	mF_Mpc_b_Ac: ARRAY[0..731] OF LREAL := [-0.00028473180920350741, -0.00064838280152378558, -0.0010871186383875045, -0.0015972149310527575, -0.0021750553811336337, -0.0028171299154482626, -0.0035200328169797839, -0.00428046085366274, -0.0050952114066324721, -0.0059611805995021831, -0.0068753614301614151, -0.0078348419065206853, -0.00883680318755997, -0.0098785177309735454, -0.010957347448640358, -0.012070741871087625, -0.013216236322055611, -0.014391450104213641, -0.015594084697021157, -0.016821921967673122, -0.018072822396016243, -0.019344723314271256, -0.02063563716234695, -0.021943649759483548, -0.023266918592916585, -0.024603671124207489, -0.025952203113843546, -0.027310876964667902, -0.02867812008465969, -0.030052423269545051, -0.031432339105682078, -0.032816480393626085, -0.034203518592746424, -0.035592182287232092, -0.036981255673790715, -0.038369577071313908, -0.039756037452751761, -0.041139578999410086, -0.042519193677855886, -0.043893921839589789, -0.04526285084361819, -0.046625113702033094, -0.047979887748683912, -0.049326393331002638, -0.050663892525022049, -0.051991687873605683, -0.053309121147888459, -0.054615572131907646, -0.055910457430385821, -0.057193229299610078, -0.058463374501335187, -0.05972041317962274, -0.06096389776051344, -0.062193411874415308, -0.063408569301077411, -0.0646090129370057, -0.065794413785165692, -0.066964469966805218, -0.068118905755219825, -0.069257470631273188, -0.070379938360475486, -0.071486106091413787, -0.072575793475319991, -0.073648841806554288, -0.074705113183774638, -0.075744489691556227, -0.076766872602218345, -0.077772181597610637, -0.078760354010605146, -0.079731344086035758, -0.080685122260822376, -0.081621674463012911, -0.082541001429472627, -0.08344311804194729, -0.084328052681223467, -0.085195846599106978, -0.086046553307938353, -0.08688023798736208, -0.087696976908065286, -0.088496856872199881, -0.089279974670201517, -0.090046436553718037, -0.0907963577243595, -0.091529861837982063, -0.092247080524217845, -0.0929481529209633, -0.093633225223539271, -0.094302450248236622, -0.094955987009962314, -0.0955940003137019, -0.096216660359515871, -0.096824142360788817, -0.09741662617545184, -0.0979942959499008, -0.098557339775334651, -0.099105949356240508, -0.099640319690754223, -0.10016064876262748, -0.1006671372445353, -0.10115998821245992, -0.10163940687089022, -0.10210560028857829, -0.10255877714459775, -0.10299914748445149, -0.10342692248597933, -0.10384231423481935, -0.10424553550917975, -0.10463679957368147, -0.10501631998203463, -0.105384310388316, -0.10574098436661702, -0.10608655523883639, -0.10642123591039374, -0.10674523871364502, -0.10705877525878353, -0.1073620562920138, -0.1076552915607895, -0.10793868968590982, -0.10821245804027231, -0.10847680263408387, 0.00028473180920350741, 0.00064838280152378558, 0.0010871186383875045, 0.0015972149310527575, 0.0021750553811336337, 0.0028171299154482626, 0.0035200328169797839, 0.00428046085366274, 0.0050952114066324721, 0.0059611805995021831, 0.0068753614301614151, 0.0078348419065206853, 0.00883680318755997, 0.0098785177309735454, 0.010957347448640358, 0.012070741871087625, 0.013216236322055611, 0.014391450104213641, 0.015594084697021157, 0.016821921967673122, 0.018072822396016243, 0.019344723314271256, 0.02063563716234695, 0.021943649759483548, 0.023266918592916585, 0.024603671124207489, 0.025952203113843546, 0.027310876964667902, 0.02867812008465969, 0.030052423269545051, 0.031432339105682078, 0.032816480393626085, 0.034203518592746424, 0.035592182287232092, 0.036981255673790715, 0.038369577071313908, 0.039756037452751761, 0.041139578999410086, 0.042519193677855886, 0.043893921839589789, 0.04526285084361819, 0.046625113702033094, 0.047979887748683912, 0.049326393331002638, 0.050663892525022049, 0.051991687873605683, 0.053309121147888459, 0.054615572131907646, 0.055910457430385821, 0.057193229299610078, 0.058463374501335187, 0.05972041317962274, 0.06096389776051344, 0.062193411874415308, 0.063408569301077411, 0.0646090129370057, 0.065794413785165692, 0.066964469966805218, 0.068118905755219825, 0.069257470631273188, 0.070379938360475486, 0.071486106091413787, 0.072575793475319991, 0.073648841806554288, 0.074705113183774638, 0.075744489691556227, 0.076766872602218345, 0.077772181597610637, 0.078760354010605146, 0.079731344086035758, 0.080685122260822376, 0.081621674463012911, 0.082541001429472627, 0.08344311804194729, 0.084328052681223467, 0.085195846599106978, 0.086046553307938353, 0.08688023798736208, 0.087696976908065286, 0.088496856872199881, 0.089279974670201517, 0.090046436553718037, 0.0907963577243595, 0.091529861837982063, 0.092247080524217845, 0.0929481529209633, 0.093633225223539271, 0.094302450248236622, 0.094955987009962314, 0.0955940003137019, 0.096216660359515871, 0.096824142360788817, 0.09741662617545184, 0.0979942959499008, 0.098557339775334651, 0.099105949356240508, 0.099640319690754223, 0.10016064876262748, 0.1006671372445353, 0.10115998821245992, 0.10163940687089022, 0.10210560028857829, 0.10255877714459775, 0.10299914748445149, 0.10342692248597933, 0.10384231423481935, 0.10424553550917975, 0.10463679957368147, 0.10501631998203463, 0.105384310388316, 0.10574098436661702, 0.10608655523883639, 0.10642123591039374, 0.10674523871364502, 0.10705877525878353, 0.1073620562920138, 0.1076552915607895, 0.10793868968590982, 0.10821245804027231, 0.10847680263408387, -1.0, -1.0, 1.0, 1.0, -0.0, -0.00028473180920350741, -0.00064838280152378558, -0.0010871186383875045, -0.0015972149310527575, -0.0021750553811336337, -0.0028171299154482626, -0.0035200328169797839, -0.00428046085366274, -0.0050952114066324721, -0.0059611805995021831, -0.0068753614301614151, -0.0078348419065206853, -0.00883680318755997, -0.0098785177309735454, -0.010957347448640358, -0.012070741871087625, -0.013216236322055611, -0.014391450104213641, -0.015594084697021157, -0.016821921967673122, -0.018072822396016243, -0.019344723314271256, -0.02063563716234695, -0.021943649759483548, -0.023266918592916585, -0.024603671124207489, -0.025952203113843546, -0.027310876964667902, -0.02867812008465969, -0.030052423269545051, -0.031432339105682078, -0.032816480393626085, -0.034203518592746424, -0.035592182287232092, -0.036981255673790715, -0.038369577071313908, -0.039756037452751761, -0.041139578999410086, -0.042519193677855886, -0.043893921839589789, -0.04526285084361819, -0.046625113702033094, -0.047979887748683912, -0.049326393331002638, -0.050663892525022049, -0.051991687873605683, -0.053309121147888459, -0.054615572131907646, -0.055910457430385821, -0.057193229299610078, -0.058463374501335187, -0.05972041317962274, -0.06096389776051344, -0.062193411874415308, -0.063408569301077411, -0.0646090129370057, -0.065794413785165692, -0.066964469966805218, -0.068118905755219825, -0.069257470631273188, -0.070379938360475486, -0.071486106091413787, -0.072575793475319991, -0.073648841806554288, -0.074705113183774638, -0.075744489691556227, -0.076766872602218345, -0.077772181597610637, -0.078760354010605146, -0.079731344086035758, -0.080685122260822376, -0.081621674463012911, -0.082541001429472627, -0.08344311804194729, -0.084328052681223467, -0.085195846599106978, -0.086046553307938353, -0.08688023798736208, -0.087696976908065286, -0.088496856872199881, -0.089279974670201517, -0.090046436553718037, -0.0907963577243595, -0.091529861837982063, -0.092247080524217845, -0.0929481529209633, -0.093633225223539271, -0.094302450248236622, -0.094955987009962314, -0.0955940003137019, -0.096216660359515871, -0.096824142360788817, -0.09741662617545184, -0.0979942959499008, -0.098557339775334651, -0.099105949356240508, -0.099640319690754223, -0.10016064876262748, -0.1006671372445353, -0.10115998821245992, -0.10163940687089022, -0.10210560028857829, -0.10255877714459775, -0.10299914748445149, -0.10342692248597933, -0.10384231423481935, -0.10424553550917975, -0.10463679957368147, -0.10501631998203463, -0.105384310388316, -0.10574098436661702, -0.10608655523883639, -0.10642123591039374, -0.10674523871364502, -0.10705877525878353, -0.1073620562920138, -0.1076552915607895, -0.10793868968590982, -0.10821245804027231, 0.0, 0.00028473180920350741, 0.00064838280152378558, 0.0010871186383875045, 0.0015972149310527575, 0.0021750553811336337, 0.0028171299154482626, 0.0035200328169797839, 0.00428046085366274, 0.0050952114066324721, 0.0059611805995021831, 0.0068753614301614151, 0.0078348419065206853, 0.00883680318755997, 0.0098785177309735454, 0.010957347448640358, 0.012070741871087625, 0.013216236322055611, 0.014391450104213641, 0.015594084697021157, 0.016821921967673122, 0.018072822396016243, 0.019344723314271256, 0.02063563716234695, 0.021943649759483548, 0.023266918592916585, 0.024603671124207489, 0.025952203113843546, 0.027310876964667902, 0.02867812008465969, 0.030052423269545051, 0.031432339105682078, 0.032816480393626085, 0.034203518592746424, 0.035592182287232092, 0.036981255673790715, 0.038369577071313908, 0.039756037452751761, 0.041139578999410086, 0.042519193677855886, 0.043893921839589789, 0.04526285084361819, 0.046625113702033094, 0.047979887748683912, 0.049326393331002638, 0.050663892525022049, 0.051991687873605683, 0.053309121147888459, 0.054615572131907646, 0.055910457430385821, 0.057193229299610078, 0.058463374501335187, 0.05972041317962274, 0.06096389776051344, 0.062193411874415308, 0.063408569301077411, 0.0646090129370057, 0.065794413785165692, 0.066964469966805218, 0.068118905755219825, 0.069257470631273188, 0.070379938360475486, 0.071486106091413787, 0.072575793475319991, 0.073648841806554288, 0.074705113183774638, 0.075744489691556227, 0.076766872602218345, 0.077772181597610637, 0.078760354010605146, 0.079731344086035758, 0.080685122260822376, 0.081621674463012911, 0.082541001429472627, 0.08344311804194729, 0.084328052681223467, 0.085195846599106978, 0.086046553307938353, 0.08688023798736208, 0.087696976908065286, 0.088496856872199881, 0.089279974670201517, 0.090046436553718037, 0.0907963577243595, 0.091529861837982063, 0.092247080524217845, 0.0929481529209633, 0.093633225223539271, 0.094302450248236622, 0.094955987009962314, 0.0955940003137019, 0.096216660359515871, 0.096824142360788817, 0.09741662617545184, 0.0979942959499008, 0.098557339775334651, 0.099105949356240508, 0.099640319690754223, 0.10016064876262748, 0.1006671372445353, 0.10115998821245992, 0.10163940687089022, 0.10210560028857829, 0.10255877714459775, 0.10299914748445149, 0.10342692248597933, 0.10384231423481935, 0.10424553550917975, 0.10463679957368147, 0.10501631998203463, 0.105384310388316, 0.10574098436661702, 0.10608655523883639, 0.10642123591039374, 0.10674523871364502, 0.10705877525878353, 0.1073620562920138, 0.1076552915607895, 0.10793868968590982, 0.10821245804027231, -0.0, -1.0, 0.0, 1.0, 1.0, 1.0, 1.0, 1.0, 1.0, 1.0, 1.0, 1.0, 1.0, 1.0, 1.0, 1.0, 1.0, 1.0, 1.0, 1.0, 1.0, 1.0, 1.0, 1.0, 1.0, 1.0, 1.0, 1.0, 1.0, 1.0, 1.0, 1.0, 1.0, 1.0, 1.0, 1.0, 1.0, 1.0, 1.0, 1.0, 1.0, 1.0, 1.0, 1.0, 1.0, 1.0, 1.0, 1.0, 1.0, 1.0, 1.0, 1.0, 1.0, 1.0, 1.0, 1.0, 1.0, 1.0, 1.0, 1.0, 1.0, 1.0, 1.0, 1.0, 1.0, 1.0, 1.0, 1.0, 1.0, 1.0, 1.0, 1.0, 1.0, 1.0, 1.0, 1.0, 1.0, 1.0, 1.0, 1.0, 1.0, 1.0, 1.0, 1.0, 1.0, 1.0, 1.0, 1.0, 1.0, 1.0, 1.0, 1.0, 1.0, 1.0, 1.0, 1.0, 1.0, 1.0, 1.0, 1.0, 1.0, 1.0, 1.0, 1.0, 1.0, 1.0, 1.0, 1.0, 1.0, 1.0, 1.0, 1.0, 1.0, 1.0, 1.0, 1.0, 1.0, 1.0, 1.0, 1.0, 1.0, 1.0, 1.0, 1.0, 1.0, 1.0, 1.0, 1.0, 1.0, 1.0, 1.0, 1.0, 1.0, 1.0, 1.0, 1.0, 1.0, 1.0, 1.0, 1.0, 1.0, 1.0, 1.0, 1.0, 1.0, 1.0, 1.0, 1.0, 1.0, 1.0, 1.0, 1.0, 1.0, 1.0, 1.0, 1.0, 1.0, 1.0, 1.0, 1.0, 1.0, 1.0, 1.0, 1.0, 1.0, 1.0, 1.0, 1.0, 1.0, 1.0, 1.0, 1.0, 1.0, 1.0, 1.0, 1.0, 1.0, 1.0, 1.0, 1.0, 1.0, 1.0, 1.0, 1.0, 1.0, 1.0, 1.0, 1.0, 1.0, 1.0, 1.0, 1.0, 1.0, 1.0, 1.0, 1.0, 1.0, 1.0, 1.0, 1.0, 1.0, 1.0, 1.0, 1.0, 1.0, 1.0, 1.0, 1.0, 1.0, 1.0, 1.0, 1.0, 1.0, 1.0, 1.0, 1.0, 1.0, 1.0, 1.0, 1.0, 1.0, 1.0, 1.0, 1.0, 1.0, 1.0, 1.0, 1.0, 1.0, 1.0, 1.0, 1.0, 1.0, 1.0, 1.0, 1.0, 1.0, 1.0, 1.0, 1.0, 1.0, 1.0, 1.0, 1.0, 0.0, 0.0, 0.0, 0.0];
	mF_Mpc_g_a: ARRAY[0..8] OF LREAL := [0.98951110734634373, -0.012366186463409425, 0.0, 0.036765047017224647, 0.96487287051035242, 0.0, 0.0, 0.0, 1.0];
	mF_Mpc_h_a: ARRAY[0..2] OF LREAL := [-2.5204929819596814E-5, -0.00021989087306674475, 0.0];
	mF_Mpc_b_Linv: ARRAY[0..8] OF LREAL := [0.2826092377312221, -0.660519995016864, 0.0, 0.0, 0.72476386636452717, 0.0, 0.0, 0.0, 0.003162277660168379];
	mF_Mpc_i_a: ARRAY[0..5] OF LREAL := [-1.6729314626197398E-6, -5.345511968919141E-6, 0.0, 0.0, 0.0, 0.0];
END_VAR



CASE ssMethodType OF
    SS_INITIALIZE: 
        (* SystemInitialize for Atomic SubSystem: '<Root>/mF_Mpc' *)
        (* InitializeConditions for Memory: '<S3>/Memory' *)

        FOR i := 0 TO 243 DO 
            Memory_PreviousInput[i] := FALSE;
        END_FOR;

        (* End of InitializeConditions for Memory: '<S3>/Memory' *)
        

        (* InitializeConditions for UnitDelay: '<S3>/last_mv' *)
        last_mv_DSTATE := 0.0;
        (* InitializeConditions for Memory: '<S3>/last_x' *)
        last_x_PreviousInput[0] := last_x_InitialCondition[0];
        last_x_PreviousInput[1] := last_x_InitialCondition[1];
        last_x_PreviousInput[2] := last_x_InitialCondition[2];
        (* End of SystemInitialize for SubSystem: '<Root>/mF_Mpc' *)
    SS_STEP: 
        (* Outputs for Atomic SubSystem: '<Root>/mF_Mpc' *)
        (* MATLAB Function: '<S23>/optimizer' incorporates:
         *  Memory: '<S3>/last_x' *)
        (* MATLAB Function 'MPC Controller/MPC/optimizer/optimizer': '<S24>:1' *)
        (* '<S24>:1:16' coder.extrinsic('mpcblock_optimizer_double_mex'); *)
        (* '<S24>:1:17' coder.extrinsic('mpcblock_optimizer_single_mex'); *)
        (* '<S24>:1:18' coder.extrinsic('mpcblock_refmd_double_mex'); *)
        (* '<S24>:1:19' coder.extrinsic('mpcblock_refmd_single_mex'); *)
        (* Inputs (in BlockDataType except iA) *)
        (* xk:         current state (either x[k|k-1] from built-in KF or external x[k|k]) *)
        (* '<S24>:1:23' xk = convertDataType(xk0,isDouble); *)
        (* '<S24>:1:250' if isDouble *)
        (* convert an input signal to double precision when necessary *)
        (* '<S24>:1:252' if isa(u,'double') *)
        (* '<S24>:1:253' y = u; *)
        (* old_u:      last mv (calculated by MPC) *)
        (* '<S24>:1:25' old_u = convertDataType(old_u0,isDouble); *)
        (* '<S24>:1:250' if isDouble *)
        (* convert an input signal to double precision when necessary *)
        (* '<S24>:1:252' if isa(u,'double') *)
        (* '<S24>:1:253' y = u; *)
        (* ym:         current measured output (used only with built-in KF) *)
        (* '<S24>:1:27' ym = convertDataType(ym0,isDouble); *)
        (* '<S24>:1:250' if isDouble *)
        (* convert an input signal to double precision when necessary *)
        (* '<S24>:1:252' if isa(u,'double') *)
        (* '<S24>:1:253' y = u; *)
        (* ref:        output reference *)
        (* '<S24>:1:29' ref = convertDataType(ref0,isDouble); *)
        (* '<S24>:1:250' if isDouble *)
        (* convert an input signal to double precision when necessary *)
        (* '<S24>:1:252' if isa(u,'double') *)
        (* '<S24>:1:253' y = u; *)
        (* md:         measured disturbance *)
        (* '<S24>:1:31' md = convertDataType(md0,isDouble); *)
        (* '<S24>:1:250' if isDouble *)
        (* convert an input signal to double precision when necessary *)
        (* '<S24>:1:252' if isa(u,'double') *)
        (* '<S24>:1:253' y = u; *)
        (* umin:       run-time MV bound *)
        (* '<S24>:1:33' umin = convertDataType(umin0,isDouble); *)
        (* umax:       run-time MV bound *)
        (* '<S24>:1:35' umax = convertDataType(umax0,isDouble); *)
        (* ymin:       run-time OV bound *)
        (* '<S24>:1:37' ymin = convertDataType(ymin0,isDouble); *)
        (* ymax:       run-time OV bound *)
        (* '<S24>:1:39' ymax = convertDataType(ymax0,isDouble); *)
        (* E:          run-time mixed constraints *)
        (* '<S24>:1:41' E = convertDataType(E0,isDouble); *)
        (* F:          run-time mixed constraints *)
        (* '<S24>:1:43' F = convertDataType(F0,isDouble); *)
        (* G:          run-time mixed constraints *)
        (* '<S24>:1:45' G = convertDataType(G0,isDouble); *)
        (* S:          run-time mixed constraints *)
        (* '<S24>:1:47' S = convertDataType(S0,isDouble); *)
        (* switch_in:  if it matches "enable_value", MPC is active in control *)
        (* '<S24>:1:49' switch_in = int32(switch_in0); *)
        (* ext_mv:     external last mv (actual) *)
        (* '<S24>:1:51' ext_mv = convertDataType(ext_mv0,isDouble); *)
        (* MVtarget:   MV reference *)
        (* '<S24>:1:53' MVtarget = convertDataType(MVtarget0,isDouble); *)
        (* ywt:        run-time OV weights *)
        (* '<S24>:1:55' ywt = convertDataType(ywt0,isDouble); *)
        (* uwt:        run-time MV weights *)
        (* '<S24>:1:57' uwt = convertDataType(uwt0,isDouble); *)
        (* duwt:       run-time DMV weights *)
        (* '<S24>:1:59' duwt = convertDataType(duwt0,isDouble); *)
        (* ewt:     run-time Slack weights *)
        (* '<S24>:1:61' ewt = convertDataType(ewt0,isDouble); *)
        (* iA:         logical previous active set (for warm start) *)
        (* Outputs (in BlockDataType except iAout) *)
        (* xk1:        x[k+1|k] from built-in KF *)
        (* u:          optimal MV *)
        (* cost:       optimal cost *)
        (* useq:       optimal MV sequence *)
        (* xseq:       optimal state sequence *)
        (* yseq:       optimal OV sequence *)
        (* status:     QP exit flag *)
        (* xest:       x[k|k] from built-in KF *)
        (* iAout:      logical current active set *)
        (* Parameters (constant) *)
        (* dimensions (int32):  *)
        (* nx, nxp, nup, nu, ny, degrees, p, nxQP, enable_value, Mrows, nCC, nv *)
        (* myindex, mvindex, mdindex, unindex, nxid, m, Ndis, numdis, maxdis *)
        (* MPC constants (BlockDataType):  *)
        (* Hinv, Kx, Ku1, Kut, Kr, Kv, Mlim, Mx, Mu1, Mv, utarget *)
        (* H, Linv, Ac, Wy, Wdu, Jm, SuJm, Su1, Sx, Hv, Wu, I1 *)
        (* A, C, B, D, Cid, Did, Ecc, Fcc, Scc, Gcc *)
        (* RYscale, RMDscale, xoff, Uscale, Yscale *)
        (* uoff, voff, yoff, myoff, RMVscale, Mdis, Vdis *)
        (* configurations (logical): *)
        (* isQP, CustomSolver, CustomSolverCodeGen, UseSuboptimalSolution, UseActiveSetSolver *)
        (* openloopflag, no_umin, no_umax, no_ymin, no_ymax, switch_inport, no_switch *)
        (* return_cost, return_mvseq, return_xseq, return_ovseq, isLTV *)
        (* no_ywt, no_uwt, no_duwt, no_rhoeps, no_md, no_ref, no_uref, no_mv *)
        (* CustomEstimation, no_cc, isHyb, isDouble *)
        (* ASOptions *)
        (* IPOptions  *)
        (* ADOptions *)
        (* MIQPOptions *)
        (* Parameters *)
        (* '<S24>:1:95' isSimulation = coder.target('Sfun') && ~coder.target('RtwForRapid') && ~coder.target('RtwForSim'); *)
        (* '<S24>:1:96' isAdaptive = false; *)
        (* '<S24>:1:97' isLTV = false; *)
        (* '<S24>:1:98' ZERO = zeros('like',ref); *)
        (* '<S24>:1:99' ONE = ones('like',ref); *)
        (* '<S24>:1:100' hasMD = nv>int32(1); *)
        (* Pre-allocate all the MEX block outputs for the simulation mode *)
        (* '<S24>:1:105' if isSimulation *)
        (* Get reference and MD signals -- accounting for previewing *)
        (* '<S24>:1:119' if isSimulation *)
        (* '<S24>:1:126' else *)
        (* When doing code generation, use M code directly *)
        (* '<S24>:1:128' [rseq, vseq, v] = mpcblock_refmd(ref,md,nv,ny,p,yoff,voff,no_md,no_ref,openloopflag, RYscale, RMDscale); *)
        i0_mpcblock_refmd(ref := flowSetpoint, md := pressureDifference, b_yoff := mF_Mpc_yoff, b_voff := mF_Mpc_voff, b_RYscale := mF_Mpc_RYscale, b_RMDscale := mF_Mpc_RMDscale);
        rseq := i0_mpcblock_refmd.rseq;
        vseq := i0_mpcblock_refmd.vseq;
        v := i0_mpcblock_refmd.v;
        (* External MV override.   *)
        (* NOTE: old_u and ext_mv input signals are dimensionless but include offset *)
        (* '<S24>:1:133' old_u = old_u - uoff; *)
        (* '<S24>:1:134' if no_mv *)
        (* '<S24>:1:135' delmv = zeros(nu,1,'like',ref); *)
        (* Obtain x[k|k] *)
        (* '<S24>:1:143' xk = xk - xoff; *)
        (* Remove offset *)
        (* '<S24>:1:144' if CustomEstimation *)
        (* '<S24>:1:147' else *)
        (* Default state estimation.     *)
        (* Scale measured output and remove offset. *)
        (* '<S24>:1:150' ym = ym.*RYscale(myindex) - myoff; *)
        (* Correct x(k|k-1) for possible external mv override. *)
        (* NOTE:  Offset was removed from x[k|k-1] at k=0. *)
        (* '<S24>:1:153' xk = xk + Bu*delmv; *)
        (* Measurement upate to x(k|k) *)
        (* '<S24>:1:155' ym_est = C(myindex,:)*xk + Dv(myindex,:)*v; *)
        (* '<S24>:1:156' y_innov = ym - ym_est; *)
        xk_idx_0 := last_x_PreviousInput[0];
        xk_idx_1 := last_x_PreviousInput[1];
        xk := last_x_PreviousInput[2];
        y_innov := (flowCurrent - mF_Mpc_myoff) - (((-10.21900021533747 * last_x_PreviousInput[0]) + (-0.12352775524810869 * last_x_PreviousInput[1])) + last_x_PreviousInput[2]);
        (* '<S24>:1:157' xest = xk + M*y_innov; *)
        rtb_xest[0] := (-6.1536996887046058E-9 * y_innov) + last_x_PreviousInput[0];
        rtb_xest[1] := (-1.4963729164443884E-7 * y_innov) + last_x_PreviousInput[1];
        rtb_xest_tmp := 0.61803395236056324 * y_innov;
        rtb_xest[2] := rtb_xest_tmp + last_x_PreviousInput[2];
        (* End of Outputs for SubSystem: '<Root>/mF_Mpc' *)
        (* Real-time MV target override *)
        (* Note: utargetValue is a vector length p*nu.   *)
        (* '<S24>:1:162' if no_uref *)
        (* no external utarget *)
        (* '<S24>:1:164' utargetValue = utarget; *)
        (* Real-time custom constraint override (scaled E/F/S) *)
        (* '<S24>:1:173' if ~no_cc *)
        (* '<S24>:1:182' return_sequence = return_mvseq || return_xseq || return_ovseq; *)
        (* '<S24>:1:183' if isSimulation *)
        (* '<S24>:1:214' else *)
        (* When doing code generation, use M code directly *)
        (* '<S24>:1:216' [u, cost, useq, status, iAout] = mpcblock_optimizer(... *)
        (* '<S24>:1:217'             rseq, vseq, umin, umax, ymin, ymax, switch_in, xest, old_u, iA, ... *)
        (* '<S24>:1:218'             isQP, nu, ny, degrees, Hinv, Kx, Ku1, Kut, Kr, Kv, Mlim, ... *)
        (* '<S24>:1:219'             Mx, Mu1, Mv, utargetValue, p, uoff, voff, yoff, ... *)
        (* '<S24>:1:220'             false, CustomSolverCodeGen, UseSuboptimalSolution, ... *)
        (* '<S24>:1:221'             UseActiveSetSolver, ASOptions, IPOptions, ADOptions, MIQPOptions, nxQP, openloopflag, ... *)
        (* '<S24>:1:222'             no_umin, no_umax, no_ymin, no_ymax, no_cc, switch_inport, ... *)
        (* '<S24>:1:223'             no_switch, enable_value, return_cost, H, return_sequence, Linv, Ac, ... *)
        (* '<S24>:1:224'             ywt, uwt, duwt, ewt, no_ywt, no_uwt, no_duwt, no_rhoeps,... *)
        (* '<S24>:1:225'             Wy, Wdu, Jm, SuJm, Su1, Sx, Hv, Wu, I1, ... *)
        (* '<S24>:1:226'             isAdaptive, isLTV, A, Bu, Bv, C, Dv, ... *)
        (* '<S24>:1:227'             Mrows, nCC, Ecc, Fcc, Scc, Gcc, RYscale, RMVscale, m, ... *)
        (* '<S24>:1:228'             isHyb, Mdis, Ndis, Vdis, numdis, maxdis); *)
        (* Outputs for Atomic SubSystem: '<Root>/mF_Mpc' *)
        (* MATLAB Function: '<S23>/optimizer' *)
        (* End of Outputs for SubSystem: '<Root>/mF_Mpc' *)
        (* Outputs for Atomic SubSystem: '<Root>/mF_Mpc' *)
        (* MATLAB Function: '<S23>/optimizer' incorporates:
         *  Memory: '<S3>/Memory'
         *  UnitDelay: '<S3>/last_mv' *)
        rMin := rtb_xest[1];
        Xnorm0 := rtb_xest[0];
        cMin := rtb_xest[2];

        FOR i := 0 TO 243 DO 
            rtb_iAout[i] := Memory_PreviousInput[i];
            a_1[i] := ((((mF_Mpc_d_a[i + 244] * rMin) + (mF_Mpc_d_a[i] * Xnorm0)) + (mF_Mpc_d_a[i + 488] * cMin)) + mF_Mpc_b_Mlim[i]) + (mF_Mpc_e_a[i] * last_mv_DSTATE);
            cTol[i] := 0.0;
        END_FOR;


        FOR k_k := 0 TO 241 DO 
            cMin := vseq[k_k];

            FOR i := 0 TO 243 DO 
                cTol[i] := (mF_Mpc_f_a[(244 * k_k) + i] * cMin) + cTol[i];
            END_FOR;

        END_FOR;

        (* End of Outputs for SubSystem: '<Root>/mF_Mpc' *)
        (* Outputs for Atomic SubSystem: '<Root>/mF_Mpc' *)
        (* MATLAB Function: '<S23>/optimizer' incorporates:
         *  UnitDelay: '<S3>/last_mv' *)

        FOR k_k := 0 TO 243 DO 
            b[k_k] :=  -(a_1[k_k] + cTol[k_k]);
        END_FOR;

        z[0] := 0.0;
        z[1] := 0.0;

        FOR i := 0 TO 1 DO 
            rMin := 0.0;

            FOR k_k := 0 TO 119 DO 
                rMin := (mF_Mpc_b_Kr[(120 * i) + k_k] * rseq[k_k]) + rMin;
            END_FOR;

            Xnorm0 := 0.0;

            FOR k_k := 0 TO 241 DO 
                Xnorm0 := (mF_Mpc_b_Kv[(242 * i) + k_k] * vseq[k_k]) + Xnorm0;
            END_FOR;

            z[i] := (((((mF_Mpc_b_Kx[(3 * i) + 1] * rtb_xest[1]) + (mF_Mpc_b_Kx[3 * i] * rtb_xest[0])) + (mF_Mpc_b_Kx[(3 * i) + 2] * rtb_xest[2])) + rMin) + (((-0.10984534103033639 * DINT_TO_LREAL(i)) + 11.520662026714231) * last_mv_DSTATE)) + Xnorm0;
        END_FOR;

        rtb_xest[0] := 0.0;
        rtb_xest[1] := 0.0;
        rtb_xest[2] := 0.0;
        i := 1;
        b_r[0] := 0.0;
        b_r[1] := 0.0;
        b_r[2] := 0.0;
        rMin := 0.0;
        cTolComputed := FALSE;
        (* End of Outputs for SubSystem: '<Root>/mF_Mpc' *)
        (* Outputs for Atomic SubSystem: '<Root>/mF_Mpc' *)
        (* MATLAB Function: '<S23>/optimizer' incorporates:
         *  Memory: '<S3>/Memory'
         *  UnitDelay: '<S3>/last_mv' *)

        FOR kDrop := 0 TO 243 DO 
            a_1[kDrop] := 0.0;
            cTol[kDrop] := 1.0;
            iC[kDrop] := 0;
        END_FOR;

        nA := 0;

        FOR tmp := 0 TO 243 DO 

            IF Memory_PreviousInput[tmp] THEN 
                nA := nA + 1;
                iC[nA - 1] := tmp + 1;
            END_IF;

        END_FOR;

        temp1 := FALSE;

        IF nA > 0 THEN 

            FOR kDrop := 0 TO 5 DO 
                Opt[kDrop] := 0.0;
            END_FOR;

            Rhs[0] := z[0];
            Rhs[3] := 0.0;
            Rhs[1] := z[1];
            Rhs[4] := 0.0;
            Rhs[2] := 0.0;
            Rhs[5] := 0.0;
            DualFeasible := FALSE;
            Xnorm0 := 0.3 * DINT_TO_LREAL(nA);

            IF Xnorm0 >= 0.5 THEN 
                tmp := TRUNC(rt_floord(u := Xnorm0 + 0.5));
            ELSE 
                tmp := 0;
            END_IF;


            IF tmp <= 5 THEN 
                tmp := 5;
            END_IF;

            ColdReset := FALSE;
            REPEAT 
                exitg3 := 0;

                IF (( NOT DualFeasible) AND (nA > 0)) AND (i <= 988) THEN 
                    kDrop := 1;

                    FOR k_k := 0 TO 8 DO 
                        RLinv[k_k] := 0.0;
                    END_FOR;

                    iSave := 0;
                    WHILE iSave <= (nA - 1) DO
                        iC_0 := iC[iSave];
                        RLinv[3 * iSave] := 0.0;
                        RLinv_tmp := (3 * iSave) + 1;
                        RLinv[RLinv_tmp] := 0.0;
                        RLinv_tmp_0 := (3 * iSave) + 2;
                        RLinv[RLinv_tmp_0] := 0.0;

                        FOR k_k := 0 TO 2 DO 
                            cMin := mF_Mpc_b_Ac[((244 * k_k) + iC_0) - 1];
                            RLinv[3 * iSave] := (mF_Mpc_b_Linv[3 * k_k] * cMin) + RLinv[3 * iSave];
                            RLinv[RLinv_tmp] := (mF_Mpc_b_Linv[(3 * k_k) + 1] * cMin) + RLinv[RLinv_tmp];
                            RLinv[RLinv_tmp_0] := (mF_Mpc_b_Linv[(3 * k_k) + 2] * cMin) + RLinv[RLinv_tmp_0];
                        END_FOR;

                        iSave := iSave + 1;
                    END_WHILE;
                    i0_qr(b_A := RLinv);
                    QQ := i0_qr.Q;
                    RR := i0_qr.b_R;
                    iSave := 0;
                    REPEAT 
                        exitg4 := 0;

                        IF iSave <= (nA - 1) THEN 

                            IF ABS(RR[(3 * iSave) + iSave]) < 1.0E-12 THEN 
                                kDrop := -2;
                                exitg4 := 1;
                            ELSE 
                                iSave := iSave + 1;
                            END_IF;

                        ELSE 

                            FOR iSave := 0 TO 2 DO 
                                cMin := mF_Mpc_b_Linv[(3 * iSave) + 1];
                                cVal := mF_Mpc_b_Linv[3 * iSave];
                                t := mF_Mpc_b_Linv[(3 * iSave) + 2];

                                FOR v_i := 0 TO 2 DO 
                                    TL[iSave + (3 * v_i)] := ((cMin * QQ[(3 * v_i) + 1]) + (cVal * QQ[3 * v_i])) + (t * QQ[(3 * v_i) + 2]);
                                END_FOR;

                            END_FOR;


                            FOR k_k := 0 TO 8 DO 
                                RLinv[k_k] := 0.0;
                            END_FOR;

                            iSave := nA - 1;
                            WHILE (iSave + 1) > 0 DO
                                RLinv_tmp := iSave + (3 * iSave);
                                RLinv[RLinv_tmp] := 1.0;
                                v_i := iSave;
                                WHILE (v_i + 1) <= nA DO
                                    RLinv_tmp_0 := (3 * v_i) + iSave;
                                    RLinv[RLinv_tmp_0] := RLinv[RLinv_tmp_0] / RR[RLinv_tmp];
                                    v_i := v_i + 1;
                                END_WHILE;

                                IF (iSave + 1) > 1 THEN 
                                    v_i := 0;
                                    WHILE v_i <= (iSave - 1) DO
                                        k_k := iSave;
                                        WHILE (k_k + 1) <= nA DO
                                            RLinv_tmp := (3 * k_k) + v_i;
                                            RLinv[RLinv_tmp] := RLinv[RLinv_tmp] - (RR[(3 * iSave) + v_i] * RLinv[(3 * k_k) + iSave]);
                                            k_k := k_k + 1;
                                        END_WHILE;
                                        v_i := v_i + 1;
                                    END_WHILE;
                                END_IF;

                                iSave := iSave - 1;
                            END_WHILE;
                            v_i := 0;
                            WHILE (v_i + 1) <= mF_Mpc_degrees DO
                                b_H[3 * v_i] := 0.0;
                                k_k := nA;
                                WHILE (k_k + 1) <= mF_Mpc_degrees DO
                                    b_H[3 * v_i] := b_H[3 * v_i] - (TL[(3 * k_k) + v_i] * TL[3 * k_k]);
                                    k_k := k_k + 1;
                                END_WHILE;
                                b_H[v_i] := b_H[3 * v_i];
                                v_i := v_i + 1;
                            END_WHILE;
                            v_i := 1;
                            WHILE (v_i + 1) <= mF_Mpc_degrees DO
                                iSave := (3 * v_i) + 1;
                                b_H[iSave] := 0.0;
                                k_k := nA;
                                WHILE (k_k + 1) <= mF_Mpc_degrees DO
                                    b_H[iSave] := b_H[iSave] - (TL[(3 * k_k) + 1] * TL[(3 * k_k) + v_i]);
                                    k_k := k_k + 1;
                                END_WHILE;
                                b_H[v_i + 3] := b_H[iSave];
                                v_i := v_i + 1;
                            END_WHILE;
                            v_i := 2;
                            WHILE (v_i + 1) <= mF_Mpc_degrees DO
                                iSave := (3 * v_i) + 2;
                                b_H[iSave] := 0.0;
                                k_k := nA;
                                WHILE (k_k + 1) <= mF_Mpc_degrees DO
                                    b_H[iSave] := b_H[iSave] - (TL[(3 * k_k) + 2] * TL[(3 * k_k) + v_i]);
                                    k_k := k_k + 1;
                                END_WHILE;
                                b_H[v_i + 6] := b_H[iSave];
                                v_i := v_i + 1;
                            END_WHILE;
                            iSave := 0;
                            WHILE iSave <= (nA - 1) DO
                                b_D[3 * iSave] := 0.0;
                                k_k := iSave;
                                WHILE (k_k + 1) <= nA DO
                                    b_D[3 * iSave] := (RLinv[(3 * k_k) + iSave] * TL[3 * k_k]) + b_D[3 * iSave];
                                    k_k := k_k + 1;
                                END_WHILE;
                                v_i := (3 * iSave) + 1;
                                b_D[v_i] := 0.0;
                                k_k := iSave;
                                WHILE (k_k + 1) <= nA DO
                                    b_D[v_i] := (TL[(3 * k_k) + 1] * RLinv[(3 * k_k) + iSave]) + b_D[v_i];
                                    k_k := k_k + 1;
                                END_WHILE;
                                v_i := (3 * iSave) + 2;
                                b_D[v_i] := 0.0;
                                k_k := iSave;
                                WHILE (k_k + 1) <= nA DO
                                    b_D[v_i] := (TL[(3 * k_k) + 2] * RLinv[(3 * k_k) + iSave]) + b_D[v_i];
                                    k_k := k_k + 1;
                                END_WHILE;
                                iSave := iSave + 1;
                            END_WHILE;
                            exitg4 := 1;
                        END_IF;

                    UNTIL NOT(exitg4 = 0)
                    END_REPEAT;

                    IF kDrop < 0 THEN 

                        IF ColdReset THEN 
                            i := -2;
                            exitg3 := 2;
                        ELSE 
                            nA := 0;

                            FOR kDrop := 0 TO 243 DO 
                                rtb_iAout[kDrop] := FALSE;
                                iC[kDrop] := 0;
                            END_FOR;

                            ColdReset := TRUE;
                        END_IF;

                    ELSE 
                        kDrop := 0;
                        WHILE kDrop <= (nA - 1) DO
                            Rhs[kDrop + 3] := b[iC[kDrop] - 1];
                            iSave := kDrop;
                            WHILE (iSave + 1) <= nA DO
                                k_k := iSave + (3 * kDrop);
                                b_U[k_k] := 0.0;
                                v_i := 0;
                                WHILE v_i <= (nA - 1) DO
                                    b_U[k_k] := (RLinv[(3 * v_i) + iSave] * RLinv[(3 * v_i) + kDrop]) + b_U[k_k];
                                    v_i := v_i + 1;
                                END_WHILE;
                                b_U[kDrop + (3 * iSave)] := b_U[k_k];
                                iSave := iSave + 1;
                            END_WHILE;
                            kDrop := kDrop + 1;
                        END_WHILE;

                        FOR kDrop := 0 TO 2 DO 
                            Opt[kDrop] := ((b_H[kDrop + 3] * Rhs[1]) + (b_H[kDrop] * Rhs[0])) + (b_H[kDrop + 6] * Rhs[2]);
                            iSave := 0;
                            WHILE iSave <= (nA - 1) DO
                                Opt[kDrop] := (b_D[(3 * iSave) + kDrop] * Rhs[iSave + 3]) + Opt[kDrop];
                                iSave := iSave + 1;
                            END_WHILE;
                        END_FOR;

                        kDrop := 0;
                        WHILE kDrop <= (nA - 1) DO
                            Opt[kDrop + 3] := ((b_D[(3 * kDrop) + 1] * Rhs[1]) + (b_D[3 * kDrop] * Rhs[0])) + (b_D[(3 * kDrop) + 2] * Rhs[2]);
                            iSave := 0;
                            WHILE iSave <= (nA - 1) DO
                                Opt[kDrop + 3] := (b_U[(3 * iSave) + kDrop] * Rhs[iSave + 3]) + Opt[kDrop + 3];
                                iSave := iSave + 1;
                            END_WHILE;
                            kDrop := kDrop + 1;
                        END_WHILE;
                        Xnorm0 := -1.0E-12;
                        kDrop := 0;
                        iSave := 3;
                        WHILE (iSave - 3) <= (nA - 1) DO
                            a_1[iC[iSave - 3] - 1] := Opt[iSave];

                            IF Opt[iSave] < Xnorm0 THEN 

                                IF (iSave - 2) <= nA THEN 
                                    kDrop := iSave - 2;
                                    Xnorm0 := Opt[iSave];
                                END_IF;

                            END_IF;

                            iSave := iSave + 1;
                        END_WHILE;

                        IF kDrop <= 0 THEN 
                            DualFeasible := TRUE;
                            rtb_xest[0] := Opt[0];
                            rtb_xest[1] := Opt[1];
                            rtb_xest[2] := Opt[2];
                        ELSE 
                            i := i + 1;

                            IF i > tmp THEN 
                                nA := 0;

                                FOR kDrop := 0 TO 243 DO 
                                    rtb_iAout[kDrop] := FALSE;
                                    iC[kDrop] := 0;
                                END_FOR;

                                ColdReset := TRUE;
                            ELSE 
                                a_1[iC[kDrop - 1] - 1] := 0.0;
                                i0_DropConstraint(kDrop := kDrop, iA := rtb_iAout, nA := nA, iC := iC);
                            END_IF;

                        END_IF;

                    END_IF;

                ELSE 

                    IF nA <= 0 THEN 

                        FOR kDrop := 0 TO 243 DO 
                            a_1[kDrop] := 0.0;
                        END_FOR;

                        cVal := z[1];
                        t := z[0];

                        FOR tmp := 0 TO 2 DO 
                            rtb_xest[tmp] := (( -mF_Mpc_b_Hinv[tmp + 3]) * cVal) + (( -mF_Mpc_b_Hinv[tmp]) * t);
                        END_FOR;

                    END_IF;

                    exitg3 := 1;
                END_IF;

            UNTIL NOT(exitg3 = 0)
            END_REPEAT;

            IF exitg3 = 1 THEN 
                temp1 := TRUE;
            END_IF;

        ELSE 
            cVal := z[1];
            t := z[0];

            FOR tmp := 0 TO 2 DO 
                rtb_xest[tmp] := (( -mF_Mpc_b_Hinv[tmp + 3]) * cVal) + (( -mF_Mpc_b_Hinv[tmp]) * t);
            END_FOR;

            temp1 := TRUE;
        END_IF;


        IF temp1 THEN 
            Xnorm0 := norm(x := rtb_xest);
            REPEAT 
                exitg2 := 0;

                IF i <= 988 THEN 
                    cMin := -1.0E-6;
                    tmp := -1;

                    FOR kDrop := 0 TO 243 DO 

                        IF  NOT cTolComputed THEN 
                            z[0] := mF_Mpc_b_Ac[kDrop] * rtb_xest[0];
                            z[1] := mF_Mpc_b_Ac[kDrop + 244] * rtb_xest[1];
                            z[2] := mF_Mpc_b_Ac[kDrop + 488] * rtb_xest[2];
                            i0_b_abs(x := z);
                            temp2 := i0_b_abs.y;
                            temp3 := maximum(x := temp2);
                            cTol[kDrop] := MAX(cTol[kDrop], temp3);
                        END_IF;


                        IF  NOT rtb_iAout[kDrop] THEN 
                            cVal := ((((mF_Mpc_b_Ac[kDrop + 244] * rtb_xest[1]) + (mF_Mpc_b_Ac[kDrop] * rtb_xest[0])) + (mF_Mpc_b_Ac[kDrop + 488] * rtb_xest[2])) - b[kDrop]) / cTol[kDrop];

                            IF cVal < cMin THEN 
                                cMin := cVal;
                                tmp := kDrop;
                            END_IF;

                        END_IF;

                    END_FOR;

                    cTolComputed := TRUE;

                    IF (tmp + 1) <= 0 THEN 
                        exitg2 := 1;
                    ELSIF i = 988 THEN 
                        i := 0;
                        exitg2 := 1;
                    ELSE 
                        REPEAT 
                            exitg1 := 0;

                            IF ((tmp + 1) > 0) AND (i <= 988) THEN 
                                temp1 := FALSE;

                                IF nA = 0 THEN 
                                    cVal := 0.0;
                                    t := 0.0;
                                    z_0 := 0.0;

                                    FOR k_k := 0 TO 2 DO 
                                        cMin := mF_Mpc_b_Ac[(244 * k_k) + tmp];
                                        cVal := (mF_Mpc_b_Hinv[3 * k_k] * cMin) + cVal;
                                        t := (mF_Mpc_b_Hinv[(3 * k_k) + 1] * cMin) + t;
                                        z_0 := (mF_Mpc_b_Hinv[(3 * k_k) + 2] * cMin) + z_0;
                                    END_FOR;

                                    z[2] := z_0;
                                    z[1] := t;
                                    z[0] := cVal;
                                    temp1 := TRUE;
                                ELSE 
                                    kDrop := 1;

                                    FOR k_k := 0 TO 8 DO 
                                        RLinv[k_k] := 0.0;
                                    END_FOR;

                                    v_i := 0;
                                    WHILE v_i <= (nA - 1) DO
                                        iC_0 := iC[v_i];
                                        RLinv[3 * v_i] := 0.0;
                                        RLinv_tmp := (3 * v_i) + 1;
                                        RLinv[RLinv_tmp] := 0.0;
                                        RLinv_tmp_0 := (3 * v_i) + 2;
                                        RLinv[RLinv_tmp_0] := 0.0;

                                        FOR k_k := 0 TO 2 DO 
                                            cMin := mF_Mpc_b_Ac[((244 * k_k) + iC_0) - 1];
                                            RLinv[3 * v_i] := (mF_Mpc_b_Linv[3 * k_k] * cMin) + RLinv[3 * v_i];
                                            RLinv[RLinv_tmp] := (mF_Mpc_b_Linv[(3 * k_k) + 1] * cMin) + RLinv[RLinv_tmp];
                                            RLinv[RLinv_tmp_0] := (mF_Mpc_b_Linv[(3 * k_k) + 2] * cMin) + RLinv[RLinv_tmp_0];
                                        END_FOR;

                                        v_i := v_i + 1;
                                    END_WHILE;
                                    i0_qr(b_A := RLinv);
                                    QQ := i0_qr.Q;
                                    RR := i0_qr.b_R;
                                    v_i := 0;
                                    REPEAT 
                                        exitg4 := 0;

                                        IF v_i <= (nA - 1) THEN 

                                            IF ABS(RR[(3 * v_i) + v_i]) < 1.0E-12 THEN 
                                                kDrop := -2;
                                                exitg4 := 1;
                                            ELSE 
                                                v_i := v_i + 1;
                                            END_IF;

                                        ELSE 

                                            FOR iSave := 0 TO 2 DO 
                                                cMin := mF_Mpc_b_Linv[(3 * iSave) + 1];
                                                cVal := mF_Mpc_b_Linv[3 * iSave];
                                                t := mF_Mpc_b_Linv[(3 * iSave) + 2];

                                                FOR v_i := 0 TO 2 DO 
                                                    TL[iSave + (3 * v_i)] := ((cMin * QQ[(3 * v_i) + 1]) + (cVal * QQ[3 * v_i])) + (t * QQ[(3 * v_i) + 2]);
                                                END_FOR;

                                            END_FOR;


                                            FOR k_k := 0 TO 8 DO 
                                                RLinv[k_k] := 0.0;
                                            END_FOR;

                                            iSave := nA - 1;
                                            WHILE (iSave + 1) > 0 DO
                                                RLinv_tmp := iSave + (3 * iSave);
                                                RLinv[RLinv_tmp] := 1.0;
                                                v_i := iSave;
                                                WHILE (v_i + 1) <= nA DO
                                                    RLinv_tmp_0 := (3 * v_i) + iSave;
                                                    RLinv[RLinv_tmp_0] := RLinv[RLinv_tmp_0] / RR[RLinv_tmp];
                                                    v_i := v_i + 1;
                                                END_WHILE;

                                                IF (iSave + 1) > 1 THEN 
                                                    v_i := 0;
                                                    WHILE v_i <= (iSave - 1) DO
                                                        k_k := iSave;
                                                        WHILE (k_k + 1) <= nA DO
                                                            RLinv_tmp := (3 * k_k) + v_i;
                                                            RLinv[RLinv_tmp] := RLinv[RLinv_tmp] - (RR[(3 * iSave) + v_i] * RLinv[(3 * k_k) + iSave]);
                                                            k_k := k_k + 1;
                                                        END_WHILE;
                                                        v_i := v_i + 1;
                                                    END_WHILE;
                                                END_IF;

                                                iSave := iSave - 1;
                                            END_WHILE;
                                            v_i := 0;
                                            WHILE (v_i + 1) <= mF_Mpc_degrees DO
                                                b_H[3 * v_i] := 0.0;
                                                k_k := nA;
                                                WHILE (k_k + 1) <= mF_Mpc_degrees DO
                                                    b_H[3 * v_i] := b_H[3 * v_i] - (TL[(3 * k_k) + v_i] * TL[3 * k_k]);
                                                    k_k := k_k + 1;
                                                END_WHILE;
                                                b_H[v_i] := b_H[3 * v_i];
                                                v_i := v_i + 1;
                                            END_WHILE;
                                            v_i := 1;
                                            WHILE (v_i + 1) <= mF_Mpc_degrees DO
                                                iSave := (3 * v_i) + 1;
                                                b_H[iSave] := 0.0;
                                                k_k := nA;
                                                WHILE (k_k + 1) <= mF_Mpc_degrees DO
                                                    b_H[iSave] := b_H[iSave] - (TL[(3 * k_k) + 1] * TL[(3 * k_k) + v_i]);
                                                    k_k := k_k + 1;
                                                END_WHILE;
                                                b_H[v_i + 3] := b_H[iSave];
                                                v_i := v_i + 1;
                                            END_WHILE;
                                            v_i := 2;
                                            WHILE (v_i + 1) <= mF_Mpc_degrees DO
                                                iSave := (3 * v_i) + 2;
                                                b_H[iSave] := 0.0;
                                                k_k := nA;
                                                WHILE (k_k + 1) <= mF_Mpc_degrees DO
                                                    b_H[iSave] := b_H[iSave] - (TL[(3 * k_k) + 2] * TL[(3 * k_k) + v_i]);
                                                    k_k := k_k + 1;
                                                END_WHILE;
                                                b_H[v_i + 6] := b_H[iSave];
                                                v_i := v_i + 1;
                                            END_WHILE;
                                            iSave := 0;
                                            WHILE iSave <= (nA - 1) DO
                                                b_D[3 * iSave] := 0.0;
                                                k_k := iSave;
                                                WHILE (k_k + 1) <= nA DO
                                                    b_D[3 * iSave] := (RLinv[(3 * k_k) + iSave] * TL[3 * k_k]) + b_D[3 * iSave];
                                                    k_k := k_k + 1;
                                                END_WHILE;
                                                v_i := (3 * iSave) + 1;
                                                b_D[v_i] := 0.0;
                                                k_k := iSave;
                                                WHILE (k_k + 1) <= nA DO
                                                    b_D[v_i] := (TL[(3 * k_k) + 1] * RLinv[(3 * k_k) + iSave]) + b_D[v_i];
                                                    k_k := k_k + 1;
                                                END_WHILE;
                                                v_i := (3 * iSave) + 2;
                                                b_D[v_i] := 0.0;
                                                k_k := iSave;
                                                WHILE (k_k + 1) <= nA DO
                                                    b_D[v_i] := (TL[(3 * k_k) + 2] * RLinv[(3 * k_k) + iSave]) + b_D[v_i];
                                                    k_k := k_k + 1;
                                                END_WHILE;
                                                iSave := iSave + 1;
                                            END_WHILE;
                                            exitg4 := 1;
                                        END_IF;

                                    UNTIL NOT(exitg4 = 0)
                                    END_REPEAT;

                                    IF kDrop <= 0 THEN 
                                        i := -2;
                                        exitg1 := 1;
                                    ELSE 

                                        FOR k_k := 0 TO 8 DO 
                                            b_U[k_k] :=  -b_H[k_k];
                                        END_FOR;

                                        cVal := 0.0;
                                        t := 0.0;
                                        z_0 := 0.0;

                                        FOR k_k := 0 TO 2 DO 
                                            cMin := mF_Mpc_b_Ac[(244 * k_k) + tmp];
                                            cVal := (b_U[3 * k_k] * cMin) + cVal;
                                            t := (b_U[(3 * k_k) + 1] * cMin) + t;
                                            z_0 := (b_U[(3 * k_k) + 2] * cMin) + z_0;
                                        END_FOR;

                                        z[2] := z_0;
                                        z[1] := t;
                                        z[0] := cVal;
                                        kDrop := 0;
                                        WHILE kDrop <= (nA - 1) DO
                                            b_r[kDrop] := ((b_D[(3 * kDrop) + 1] * mF_Mpc_b_Ac[tmp + 244]) + (b_D[3 * kDrop] * mF_Mpc_b_Ac[tmp])) + (b_D[(3 * kDrop) + 2] * mF_Mpc_b_Ac[tmp + 488]);
                                            kDrop := kDrop + 1;
                                        END_WHILE;
                                        temp1 := TRUE;
                                    END_IF;

                                END_IF;


                                IF temp1 THEN 
                                    kDrop := 0;
                                    cMin := 0.0;
                                    DualFeasible := TRUE;
                                    ColdReset := TRUE;

                                    IF nA > 0 THEN 
                                        iSave := 0;
                                        REPEAT 
                                            exitg4 := 0;

                                            IF iSave <= (nA - 1) THEN 

                                                IF b_r[iSave] >= 1.0E-12 THEN 
                                                    ColdReset := FALSE;
                                                    exitg4 := 1;
                                                ELSE 
                                                    iSave := iSave + 1;
                                                END_IF;

                                            ELSE 
                                                exitg4 := 1;
                                            END_IF;

                                        UNTIL NOT(exitg4 = 0)
                                        END_REPEAT;
                                    END_IF;


                                    IF (nA <> 0) AND ( NOT ColdReset) THEN 
                                        v_i := 0;
                                        WHILE v_i <= (nA - 1) DO

                                            IF b_r[v_i] > 1.0E-12 THEN 
                                                cVal := a_1[iC[v_i] - 1] / b_r[v_i];

                                                IF (kDrop = 0) OR (cVal < rMin) THEN 
                                                    rMin := cVal;
                                                    kDrop := v_i + 1;
                                                END_IF;

                                            END_IF;

                                            v_i := v_i + 1;
                                        END_WHILE;

                                        IF kDrop > 0 THEN 
                                            cMin := rMin;
                                            DualFeasible := FALSE;
                                        END_IF;

                                    END_IF;

                                    t := mF_Mpc_b_Ac[tmp + 244];
                                    z_0 := mF_Mpc_b_Ac[tmp + 488];
                                    cVal := ((t * z[1]) + (z[0] * mF_Mpc_b_Ac[tmp])) + (z_0 * z[2]);

                                    IF cVal <= 0.0 THEN 
                                        cVal := 0.0;
                                        ColdReset := TRUE;
                                    ELSE 
                                        cVal := (b[tmp] - (((t * rtb_xest[1]) + (mF_Mpc_b_Ac[tmp] * rtb_xest[0])) + (z_0 * rtb_xest[2]))) / cVal;
                                        ColdReset := FALSE;
                                    END_IF;


                                    IF DualFeasible AND ColdReset THEN 
                                        i := -1;
                                        exitg1 := 1;
                                    ELSE 

                                        IF ColdReset THEN 
                                            t := cMin;
                                        ELSIF DualFeasible THEN 
                                            t := cVal;
                                        ELSIF cMin < cVal THEN 
                                            t := cMin;
                                        ELSE 
                                            t := cVal;
                                        END_IF;

                                        v_i := 0;
                                        WHILE v_i <= (nA - 1) DO
                                            a_1[iC[v_i] - 1] := a_1[iC[v_i] - 1] - (t * b_r[v_i]);

                                            IF iC[v_i] <= 244 THEN 

                                                IF a_1[iC[v_i] - 1] < 0.0 THEN 
                                                    a_1[iC[v_i] - 1] := 0.0;
                                                END_IF;

                                            END_IF;

                                            v_i := v_i + 1;
                                        END_WHILE;
                                        a_1[tmp] := a_1[tmp] + t;

                                        IF ABS(t - cMin) < 2.2204460492503131E-16 THEN 
                                            i0_DropConstraint(kDrop := kDrop, iA := rtb_iAout, nA := nA, iC := iC);
                                        END_IF;


                                        IF  NOT ColdReset THEN 
                                            rtb_xest[0] := (t * z[0]) + rtb_xest[0];
                                            rtb_xest[1] := (t * z[1]) + rtb_xest[1];
                                            rtb_xest[2] := (t * z[2]) + rtb_xest[2];

                                            IF ABS(t - cVal) < 2.2204460492503131E-16 THEN 

                                                IF nA = mF_Mpc_degrees THEN 
                                                    i := -1;
                                                    exitg1 := 1;
                                                ELSE 
                                                    nA := nA + 1;
                                                    iC[nA - 1] := tmp + 1;
                                                    kDrop := nA - 1;
                                                    REPEAT 
                                                        exitg4 := 0;

                                                        IF (kDrop + 1) > 1 THEN 
                                                            k_k := iC[kDrop - 1];

                                                            IF iC[kDrop] > k_k THEN 
                                                                exitg4 := 1;
                                                            ELSE 
                                                                iSave := iC[kDrop];
                                                                iC[kDrop] := k_k;
                                                                iC[kDrop - 1] := iSave;
                                                                kDrop := kDrop - 1;
                                                            END_IF;

                                                        ELSE 
                                                            exitg4 := 1;
                                                        END_IF;

                                                    UNTIL NOT(exitg4 = 0)
                                                    END_REPEAT;
                                                    rtb_iAout[tmp] := TRUE;
                                                    tmp := -1;
                                                    i := i + 1;
                                                END_IF;

                                            ELSE 
                                                i := i + 1;
                                            END_IF;

                                        ELSE 
                                            i := i + 1;
                                        END_IF;

                                    END_IF;

                                END_IF;

                            ELSE 
                                cMin := norm(x := rtb_xest);

                                IF ABS(cMin - Xnorm0) > 0.001 THEN 
                                    Xnorm0 := cMin;
                                    i0_abs_a(x := b);
                                    temp4 := i0_abs_a.y;
                                    i0_maximum2(x := temp4, y := 1.0);
                                    cTol := i0_maximum2.ex;
                                    cTolComputed := FALSE;
                                END_IF;

                                exitg1 := 2;
                            END_IF;

                        UNTIL NOT(exitg1 = 0)
                        END_REPEAT;

                        IF exitg1 = 1 THEN 
                            exitg2 := 1;
                        END_IF;

                    END_IF;

                ELSE 
                    exitg2 := 1;
                END_IF;

            UNTIL NOT(exitg2 = 0)
            END_REPEAT;
        END_IF;


        IF (i < 0) OR (i = 0) THEN 
            rtb_xest[0] := 0.0;
        END_IF;

        Xnorm0 := last_mv_DSTATE + rtb_xest[0];
        (* End of Outputs for SubSystem: '<Root>/mF_Mpc' *)
        (* '<S24>:1:231' if return_xseq || return_ovseq *)
        (* '<S24>:1:233' else *)
        (* '<S24>:1:234' yseq = zeros(p+1,ny,'like',rseq); *)
        (* '<S24>:1:235' xseq = zeros(p+1,nxQP,'like',rseq); *)
        (* '<S24>:1:238' if CustomEstimation *)
        (* '<S24>:1:240' else *)
        (* update x[k+1|k], assuming that above u and v will be applied. *)
        (* '<S24>:1:242' xk1 = A*xk + Bu*(u - uoff) + Bv*v + L*y_innov; *)
        (* '<S24>:1:244' xk1 = xk1 + xoff; *)
        (* Updated state must include offset *)
        (* return xest in original value *)
        (* '<S24>:1:247' xest = xest + xoff; *)
        (* Outputs for Atomic SubSystem: '<Root>/mF_Mpc' *)
        (* Update for Memory: '<S3>/Memory' *)

        FOR i := 0 TO 243 DO 
            Memory_PreviousInput[i] := rtb_iAout[i];
        END_FOR;

        (* End of Update for Memory: '<S3>/Memory' *)
        

        (* Update for UnitDelay: '<S3>/last_mv' incorporates:
         *  MATLAB Function: '<S23>/optimizer' *)
        last_mv_DSTATE := Xnorm0;
        (* End of Outputs for SubSystem: '<Root>/mF_Mpc' *)
        (* Outputs for Atomic SubSystem: '<Root>/mF_Mpc' *)
        (* MATLAB Function: '<S23>/optimizer' *)

        FOR k_k := 0 TO 2 DO 
            rtb_xest[k_k] := (((mF_Mpc_g_a[k_k + 3] * xk_idx_1) + (mF_Mpc_g_a[k_k] * xk_idx_0)) + (mF_Mpc_g_a[k_k + 6] * xk)) + (mF_Mpc_h_a[k_k] * Xnorm0);
        END_FOR;

        xk := 0.0;
        rMin := 0.0;

        FOR k_k := 0 TO 1 DO 
            cMin := v[k_k];
            xk := (mF_Mpc_i_a[3 * k_k] * cMin) + xk;
            rMin := (mF_Mpc_i_a[(3 * k_k) + 1] * cMin) + rMin;
        END_FOR;

        (* End of Outputs for SubSystem: '<Root>/mF_Mpc' *)
        (* Outputs for Atomic SubSystem: '<Root>/mF_Mpc' *)
        (* Update for Memory: '<S3>/last_x' incorporates:
         *  MATLAB Function: '<S23>/optimizer' *)
        last_x_PreviousInput[0] := (rtb_xest[0] + xk) + (-1.1590576263587683E-8 * y_innov);
        last_x_PreviousInput[1] := (rtb_xest[1] + rMin) + (-1.443048653146427E-7 * y_innov);
        last_x_PreviousInput[2] := rtb_xest_tmp + rtb_xest[2];
        (* Outport: '<Root>/valveCommand' incorporates:
         *  MATLAB Function: '<S23>/optimizer' *)
        valveCommand := Xnorm0;
        (* End of Outputs for SubSystem: '<Root>/mF_Mpc' *)
END_CASE;

END_FUNCTION_BLOCK

(* stored: Version 1.1.0.1, ProductVersion 3.1.4024.9
   POU mF_Mpc: Id {c1e53d2d-0aec-4bb0-babd-278309e65bdb}, SpecialFunc None *)
